(*
SPDX-FileCopyrightText: © 2026 Oleksandr Tiutyk <trofimich@gmail.com>
SPDX-License-Identifier: MIT
License: https://opensource.org/license/mit
*)

(*!
<summary>Selects the SET_ERROR_AND_CONTINUE reaction for every exception.</summary>
<description>
Stateless policy: does not inspect or retain arguments, allocate memory or raise exceptions. The caller
applies the reaction and performs logging.
</description>
*)

{attribute 'no_explicit_call' := 'do not call this function block directly'}
FUNCTION_BLOCK SetErrorAndContinueExceptionHandlingPolicy EXTENDS Object IMPLEMENTS IExceptionHandlingPolicy
VAR_STAT
	//! <summary>Class name shared by all instances of this function block.</summary>
	{attribute 'hide'} 
	_ClassName : STRING := __POUNAME();
END_VAR

{attribute 'monitoring' := 'call'}
PROPERTY ClassName : REFERENCE TO STRING
GET
ClassName REF= _ClassName;
END_GET
END_PROPERTY

(*!
<summary>Returns SET_ERROR_AND_CONTINUE.</summary>
<description>
Only selects the reaction; does not modify the handling object or exception. Descendants cannot change this
fixed reaction; implement IExceptionHandlingPolicy separately for another policy.
</description>
*)
METHOD FINAL HandleException : EXCEPTION_REACTION
VAR_INPUT
	exception : IReadOnlyException;
	handlingObject : IObject;
END_VAR
VAR_IN_OUT CONSTANT
	failedMethodName : STRING(255);
END_VAR
HandleException := EXCEPTION_REACTION.SET_ERROR_AND_CONTINUE;
END_METHOD

(*!
<summary>Provides the library namespace used in diagnostics.</summary>
<description>
Borrowed read-only reference to the compiler-initialized library namespace; no ownership transfer.
</description>
*)
{attribute 'monitoring' := 'call'}
PROPERTY NamespaceName : REFERENCE TO STRING
GET
NamespaceName REF= CurrentNamespace.Name;
END_GET
END_PROPERTY

(*!
<summary>Reports the byte size of this concrete instance.</summary>
<description>
Uses XSIZEOF on the instance. Does not include separately allocated payloads or prove that an arbitrary
address is valid.
</description>
*)
{attribute 'monitoring' := 'call'}
PROPERTY SelfSize : ULINT
GET
SelfSize := XSIZEOF(THIS^);
END_GET
END_PROPERTY

END_FUNCTION_BLOCK

(* stored: Version 1.1.0.1
   POU SetErrorAndContinueExceptionHandlingPolicy: Id {a4eb2320-3400-4dc2-8031-b55b6e1bbfa3}, SpecialFunc None
   Property ClassName: Id {3ac1fd6a-8981-46e7-88fa-adfce8200fbf}
   Get Get: Id {e0a59f69-f2b1-4954-bbc5-f99626dcbdee}
   Method HandleException: Id {462be713-1109-4737-a605-c6d09182fca9}
   Property NamespaceName: Id {12125e62-a5f3-4101-949a-c95b577951f5}
   Get Get: Id {d53a3505-556c-4128-a9b8-62085a2d05b4}
   Property SelfSize: Id {cd0a5ef3-cdc3-45f0-afdb-f57972fae1ca}
   Get Get: Id {9eb177ce-67e4-410e-aed0-e7613e6a2b75} *)
